Fanuc KAREL source: kb00008.compact.KL

PROGRAM KB00008
%STACKSIZE=65535
%PRIORITY=65535
%NOLOCKGROUP
VAR
P1 : REAL
RESULT : REAL
BEGIN
P1=1.0
RESULT=ASIN(P1)
END KB00008
